Fanuc KAREL source: kd00031.KL

-- PROVISIONAL review KL for V1013-1; original PC SHA256 f7893b4cac1c56ea217ddf564f7c87f0238adfc490f46c66e30797fab2bc7055
-- Incomplete behavior may be omitted. Consult companion uncertainty JSON. Do not deploy.
PROGRAM KD00031
%NOLOCKGROUP
VAR
  I : INTEGER
  J : INTEGER
  B : BOOLEAN
  R : REAL
  S : STRING[80]
BEGIN
  -- UNRESOLVED_PC offsets 5-21; opcodes 9D,81,18,9C,12,22,9D,13,04
  -- UNRESOLVED_PC offsets 26-30; opcodes 7F
END KD00031
